// TIA Portal project "Anvil_works" (V20)

(* hardware
DEVICE "S7-1500/ET200MP station_1"  S7-1500 station
   slot 0: "Rail_0"  Rack  6ES7 590-1***0-0AA0
   slot 1: "PLC_1"  CPU 1511-1 PN  6ES7 511-1AK01-0AB0  V2.9
      slot 3: "CPU display_1"  6ES7591-1AA00-0AA0
      slot 32768: "PROFINET interface_1"  X1
         slot 32769: "Port_1"  X1 P1
         slot 32770: "Port_2"  X1 P2
      slot 34817: "Virtual CP interface port_1"  Virtual CP interface port  Virtual CP interface port
   slot 2: "DI 16x24VDC BA_1"  DI 16x24VDC BA  6ES7 521-1BH10-0AA0  V1.1
   slot 3: "AI 8xU/I/RTD/TC ST_1"  AI 8xU/I/RTD/TC ST  6ES7 531-7KF00-0AB0  V2.2
*)

// ===== PLC "PLC_1"  CPU 1511-1 PN =====

VAR_GLOBAL   // PLC tag table "Default tag table"
   "TempBit" AT %M0.0 : Bool;
   "furnance1Pulse" AT %I0.0 : Bool;
   "furnance2Pulse" AT %I0.1 : Bool;
   "furnance3Pulse" AT %I0.2 : Bool;
   "hardnessInput" AT %IW2 : Int;   // Hardness sensor, analog input channel 0
END_VAR

DATA_BLOCK "DB_AnvilQueue"   // DB1
{ S7_Optimized_Access := 'TRUE' }
VERSION : 0.1
   VAR
      items : Array[0..9] of Struct
         furnace : Int;
         timestamp : DTL;
         hardness : Int;
      END_STRUCT;
      readIndex : Int;
      writeIndex : Int;
      count : Int;
      furnance1PulseDetected : Bool;
      furnance2PulseDetected : Bool;
      furnance3PulseDetected : Bool;
   END_VAR
BEGIN
END_DATA_BLOCK

DATA_BLOCK "DB_AnvilProcess"   // DB2
{ S7_Optimized_Access := 'FALSE' }
VERSION : 0.1
   VAR
      hardnessSensor : Int;
      trigger : Bool;
      ready : Bool;
      done : Bool;
      fetchRequest : Bool;
      anvil : Struct
         furnace : Int;
         timestamp : DTL;
         hardness : Int;
      END_STRUCT;
      donePulse : Bool;
   END_VAR
BEGIN
END_DATA_BLOCK

FUNCTION "FC_EnqueueAnvil" : Void   // FC1, SCL
{ S7_Optimized_Access := 'TRUE' }
VERSION : 0.1
   VAR_INPUT
      Pulse : Bool;
      FurnaceID : Int;
   END_VAR
   VAR_OUTPUT
      Added : Bool;
      QueueFull : Bool;
      Error : Bool;
   END_VAR
   VAR_TEMP
      Now : DTL;
      ClockStatus : Int;
   END_VAR
BEGIN
   #Added := FALSE;
   #QueueFull := FALSE;
   #Error := FALSE;

   IF #Pulse THEN
       IF (#FurnaceID < 1) OR (#FurnaceID > 3) THEN
           #Error := TRUE;

       ELSIF "DB_AnvilQueue".count >= 10 THEN
           #QueueFull := TRUE;

       ELSIF ("DB_AnvilQueue".writeIndex < 0)
           OR ("DB_AnvilQueue".writeIndex > 9)
           OR ("DB_AnvilQueue".count < 0) THEN
           #Error := TRUE;

       ELSE
           #ClockStatus := RD_SYS_T(OUT => #Now);

           IF #ClockStatus = 0 THEN
               "DB_AnvilQueue".items["DB_AnvilQueue".writeIndex].furnace := #FurnaceID;
               "DB_AnvilQueue".items["DB_AnvilQueue".writeIndex].timestamp := #Now;
               "DB_AnvilQueue".items["DB_AnvilQueue".writeIndex].hardness := "DB_AnvilProcess".hardnessSensor;

               "DB_AnvilQueue".writeIndex :=
               "DB_AnvilQueue".writeIndex + 1;

               IF "DB_AnvilQueue".writeIndex >= 10 THEN
                   "DB_AnvilQueue".writeIndex := 0;
               END_IF;

               "DB_AnvilQueue".count :=
               "DB_AnvilQueue".count + 1;

               #Added := TRUE;

           ELSE
               #Error := TRUE;
           END_IF;

       END_IF;

   END_IF;
END_FUNCTION

ORGANIZATION_BLOCK "Main"   // OB1, LAD, ProgramCycle
TITLE = "Main Program Sweep (Cycle)"
{ S7_Optimized_Access := 'TRUE' }
VERSION : 0.1
   VAR_INPUT
      Initial_Call : Bool;   // Initial call of this OB
      Remanence : Bool;   // =True, if remanent data are available
   END_VAR
   VAR_TEMP
      Temp_Added : Bool;
      Temp_QueueFull : Bool;
      Temp_Error : Bool;
   END_VAR
BEGIN

REGION Network 1: Leitura da fila e ativação do Ready
   // Verifica se existem bigornas disponíveis (Count > 0). Copia a bigorna da posição ReadIndex para a estrutura Anvil e ativa o sinal Ready.
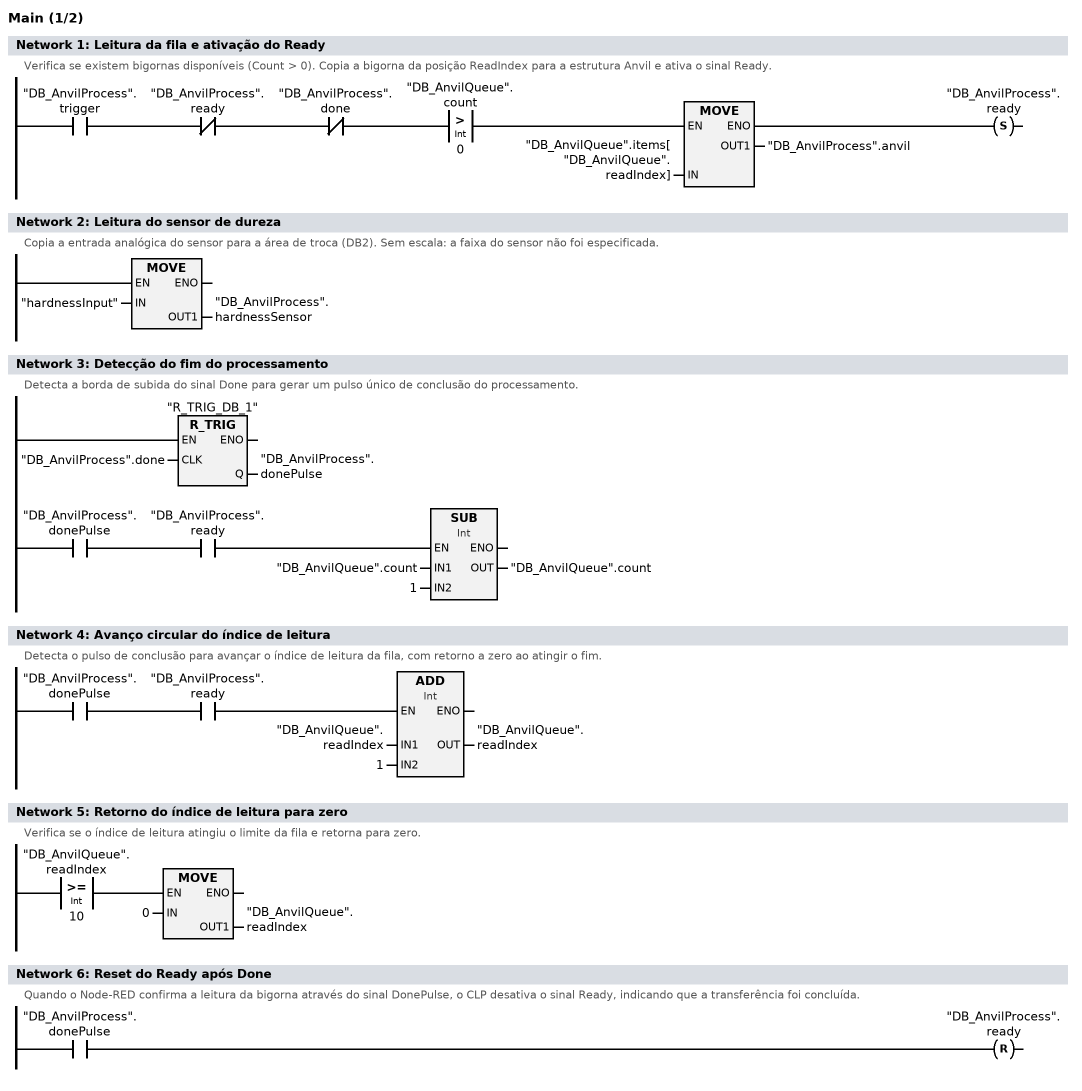
   RUNG wire#powerrail
      Contact( "DB_AnvilProcess".trigger )
      I_Contact( "DB_AnvilProcess".ready )
      I_Contact( "DB_AnvilProcess".done )
      { S7_Templates := "SrcType := Int" } GT_Contact(in1 := "DB_AnvilQueue".count, in2 := 0)
      Move(in := "DB_AnvilQueue".items["DB_AnvilQueue".readIndex], out1 => "DB_AnvilProcess".anvil)
      S_Coil( "DB_AnvilProcess".ready )
   END_RUNG
   // the same network as SCL:
   IF "DB_AnvilProcess".trigger AND NOT "DB_AnvilProcess".ready AND NOT "DB_AnvilProcess".done AND ("DB_AnvilQueue".count > 0) THEN
       "DB_AnvilProcess".anvil := "DB_AnvilQueue".items["DB_AnvilQueue".readIndex];
       "DB_AnvilProcess".ready := TRUE;
   END_IF;
END_REGION

REGION Network 2: Leitura do sensor de dureza
   // Copia a entrada analógica do sensor para a área de troca (DB2). Sem escala: a faixa do sensor não foi especificada.
   RUNG wire#powerrail
      Move(in := "hardnessInput", out1 => "DB_AnvilProcess".hardnessSensor)
   END_RUNG
   // the same network as SCL:
   "DB_AnvilProcess".hardnessSensor := "hardnessInput";
END_REGION

REGION Network 3: Detecção do fim do processamento
   // Detecta a borda de subida do sinal Done para gerar um pulso único de conclusão do processamento.
   "R_TRIG_DB_1"(CLK := "DB_AnvilProcess".done, Q => "DB_AnvilProcess".donePulse);   // R_TRIG
   IF "DB_AnvilProcess".donePulse AND "DB_AnvilProcess".ready THEN
       "DB_AnvilQueue".count := "DB_AnvilQueue".count - 1;
   END_IF;
END_REGION

REGION Network 4: Avanço circular do índice de leitura
   // Detecta o pulso de conclusão para avançar o índice de leitura da fila, com retorno a zero ao atingir o fim.
   RUNG wire#powerrail
      Contact( "DB_AnvilProcess".donePulse )
      Contact( "DB_AnvilProcess".ready )
      { S7_Templates := "SrcType := Int" } Add(in1 := "DB_AnvilQueue".readIndex, in2 := 1, out => "DB_AnvilQueue".readIndex)
   END_RUNG
   // the same network as SCL:
   IF "DB_AnvilProcess".donePulse AND "DB_AnvilProcess".ready THEN
       "DB_AnvilQueue".readIndex := "DB_AnvilQueue".readIndex + 1;
   END_IF;
END_REGION

REGION Network 5: Retorno do índice de leitura para zero
   // Verifica se o índice de leitura atingiu o limite da fila e retorna para zero.
   RUNG wire#powerrail
      { S7_Templates := "SrcType := Int" } GE_Contact(in1 := "DB_AnvilQueue".readIndex, in2 := 10)
      Move(in := 0, out1 => "DB_AnvilQueue".readIndex)
   END_RUNG
   // the same network as SCL:
   IF "DB_AnvilQueue".readIndex >= 10 THEN "DB_AnvilQueue".readIndex := 0; END_IF;
END_REGION

REGION Network 6: Reset do Ready após Done
   // Quando o Node-RED confirma a leitura da bigorna através do sinal DonePulse, o CLP desativa o sinal Ready, indicando que a transferência foi concluída.
   RUNG wire#powerrail
      Contact( "DB_AnvilProcess".donePulse )
      R_Coil( "DB_AnvilProcess".ready )
   END_RUNG
   // the same network as SCL:
   IF "DB_AnvilProcess".donePulse THEN "DB_AnvilProcess".ready := FALSE; END_IF;
END_REGION

REGION Network 7: Limpeza dos dados da bigorna
   // Quando o DonePulse ativa, limpa os dados da bigorna.
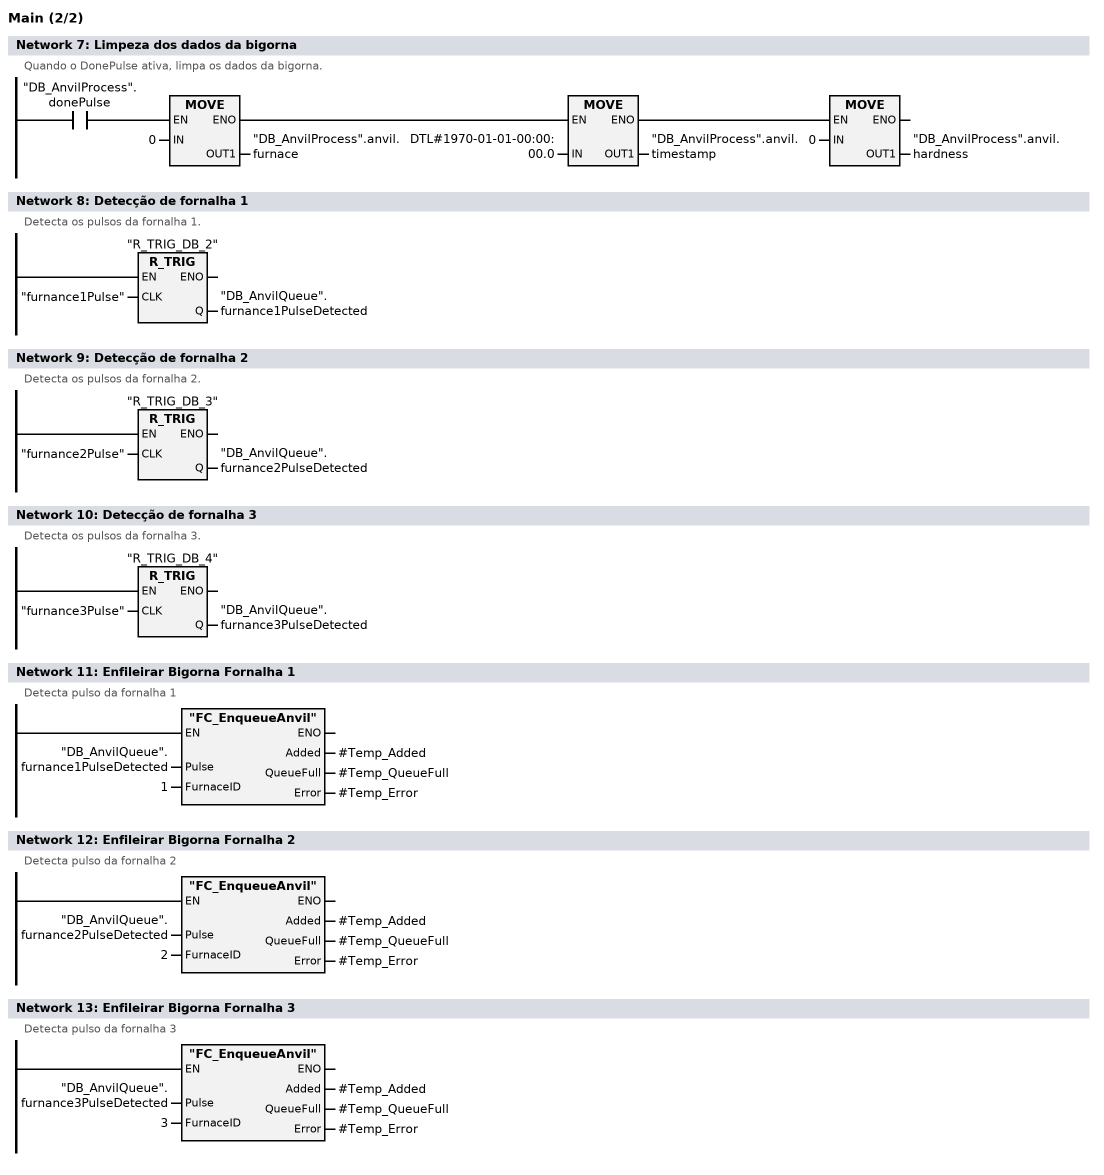
   RUNG wire#powerrail
      Contact( "DB_AnvilProcess".donePulse )
      Move(in := 0, out1 => "DB_AnvilProcess".anvil.furnace)
      Move(in := DTL#1970-01-01-00:00:00.0, out1 => "DB_AnvilProcess".anvil.timestamp)
      Move(in := 0, out1 => "DB_AnvilProcess".anvil.hardness)
   END_RUNG
   // the same network as SCL:
   IF "DB_AnvilProcess".donePulse THEN
       "DB_AnvilProcess".anvil.furnace := 0;
       "DB_AnvilProcess".anvil.timestamp := DTL#1970-01-01-00:00:00.0;
       "DB_AnvilProcess".anvil.hardness := 0;
   END_IF;
END_REGION

REGION Network 8: Detecção de fornalha 1
   // Detecta os pulsos da fornalha 1.
   "R_TRIG_DB_2"(CLK := "furnance1Pulse", Q => "DB_AnvilQueue".furnance1PulseDetected);   // R_TRIG
END_REGION

REGION Network 9: Detecção de fornalha 2
   // Detecta os pulsos da fornalha 2.
   "R_TRIG_DB_3"(CLK := "furnance2Pulse", Q => "DB_AnvilQueue".furnance2PulseDetected);   // R_TRIG
END_REGION

REGION Network 10: Detecção de fornalha 3
   // Detecta os pulsos da fornalha 3.
   "R_TRIG_DB_4"(CLK := "furnance3Pulse", Q => "DB_AnvilQueue".furnance3PulseDetected);   // R_TRIG
END_REGION

REGION Network 11: Enfileirar Bigorna Fornalha 1
   // Detecta pulso da fornalha 1
   RUNG wire#powerrail
      "FC_EnqueueAnvil"(Pulse := "DB_AnvilQueue".furnance1PulseDetected, FurnaceID := 1, Added => #Temp_Added, QueueFull => #Temp_QueueFull, Error => #Temp_Error)
   END_RUNG
   // the same network as SCL:
   "FC_EnqueueAnvil"(Pulse := "DB_AnvilQueue".furnance1PulseDetected,
                     FurnaceID := 1,
                     Added => #Temp_Added,
                     QueueFull => #Temp_QueueFull,
                     Error => #Temp_Error);
END_REGION

REGION Network 12: Enfileirar Bigorna Fornalha 2
   // Detecta pulso da fornalha 2
   RUNG wire#powerrail
      "FC_EnqueueAnvil"(Pulse := "DB_AnvilQueue".furnance2PulseDetected, FurnaceID := 2, Added => #Temp_Added, QueueFull => #Temp_QueueFull, Error => #Temp_Error)
   END_RUNG
   // the same network as SCL:
   "FC_EnqueueAnvil"(Pulse := "DB_AnvilQueue".furnance2PulseDetected,
                     FurnaceID := 2,
                     Added => #Temp_Added,
                     QueueFull => #Temp_QueueFull,
                     Error => #Temp_Error);
END_REGION

REGION Network 13: Enfileirar Bigorna Fornalha 3
   // Detecta pulso da fornalha 3
   RUNG wire#powerrail
      "FC_EnqueueAnvil"(Pulse := "DB_AnvilQueue".furnance3PulseDetected, FurnaceID := 3, Added => #Temp_Added, QueueFull => #Temp_QueueFull, Error => #Temp_Error)
   END_RUNG
   // the same network as SCL:
   "FC_EnqueueAnvil"(Pulse := "DB_AnvilQueue".furnance3PulseDetected,
                     FurnaceID := 3,
                     Added => #Temp_Added,
                     QueueFull => #Temp_QueueFull,
                     Error => #Temp_Error);
END_REGION
END_ORGANIZATION_BLOCK